RoboDK station: PICK1.rdk

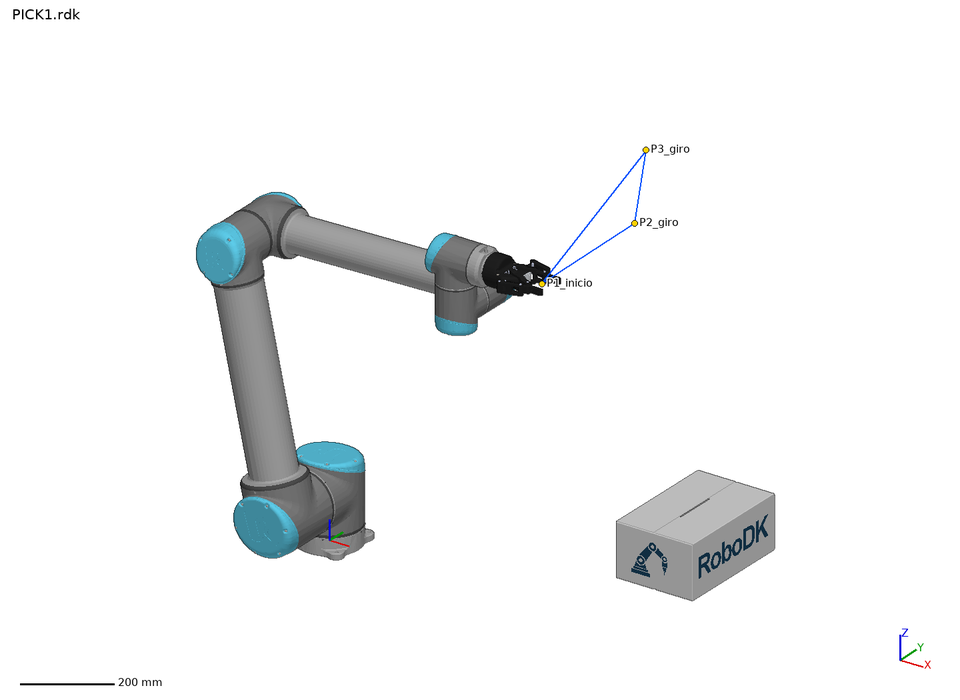
[picture v0: the station drawn from its stored meshes, robots at their saved joint values, targets as dots, program paths as lines]
Station Nueva Estación (1) (saved by RoboDK 6.1.1). Poses are relative to the parent item; angles as X-Y-Z fixed-axis rotations.
  - frame UR10 Base at (0, 0, 0) mm
    - robot UR10: 6 axes, payload 10 kg, reach 1300 mm, repeatability 0.1 mm, weight 28.9 kg
        modified DH rows (alpha deg, a mm, theta deg, d mm): 0, 0, 0, 128; 90, 0, 180, 0; 0, 612.7, 0, 0; 0, 571.6, 0, 163.9; -90, 0, 0, 115.7; 90, 0, 180, 92.2
        joint limits [-360, -360, -360, -360, -360, -360] to [360, 360, 360, 360, 360, 360]; home [0, -90, -90, 0, 90, 0]; saved at [0, -77.766, -100.839, -1.395, 90, 0]
      - tool RobotiQ 2F-85 Gripper (Closed), TCP at (0, 0, 130) mm, size 134.4 x 75 x 157.6 mm
    - target P1_inicio (Cartesian target) at (663.8, -163.9, 856.4) mm, rotated rx -90 ry 0 rz -90 deg; joints [0, -90, -90, 0, 90, 0] of UR10
    - target P2_giro (Cartesian target) at (656.82, 189.96, 856.4) mm, rotated rx -90 ry 0 rz -60 deg; joints [30, -90, -90, 0, 90, 0] of UR10
    - target P3_giro (Cartesian target) at (473.84, 492.92, 856.4) mm, rotated rx -90 ry 0 rz -30 deg; joints [60, -90, -90, 0, 90, 0] of UR10
    - object Caja at (600, 200, 0) mm, size 199 x 305.1 x 133.7 mm, geometry from Box-12x7in-Closed.sld
  - program Secuencia_UR10 (6 instructions, listed below)
  - Python program Prog2 (listed below)
  - Python program Prog3 (listed below)
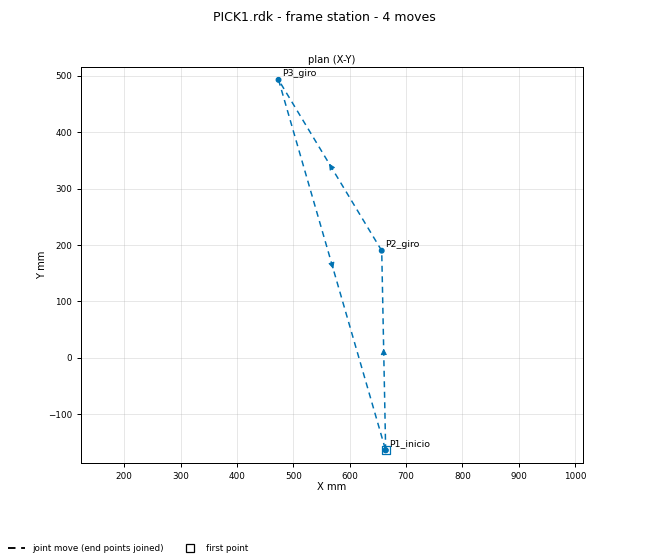
[picture p0: tool path of PICK1.rdk in frame station, 4 of 4 moves have a stored position in this frame; points joined in program order, loops and branches not executed]

--- program Secuencia_UR10 (robot UR10) ---
  Est. Ref.: UR10 Base
  MoveJ (P1_inicio)
  MoveJ (P2_giro)
  MoveJ (P3_giro)
  MoveJ (P1_inicio)
  Establecer velocidad (500.0 mm/s)

--- Python program Prog2 ---
from robodk.robolink import *

RDK = Robolink()

robot = RDK.Item('UR10', ITEM_TYPE_ROBOT)

p1 = RDK.Item('P1_inicio', ITEM_TYPE_TARGET)
p2 = RDK.Item('P2_giro', ITEM_TYPE_TARGET)
p3 = RDK.Item('P3_giro', ITEM_TYPE_TARGET)

# Verificar que existan los elementos
if not all(item.Valid() for item in [robot, p1, p2, p3]):
    raise Exception("No se encontro el robot o algun punto")

# Velocidad articular
robot.setSpeedJoints(20)

# Secuencia del brazo robotico
robot.MoveJ(p1)
robot.MoveJ(p2)
robot.MoveJ(p3)
robot.MoveJ(p1)

print("Secuencia completada")

--- Python program Prog3 ---
# -*- coding: utf-8 -*-
# Pick & Place UR10 + Robotiq 2F-85 en RoboDK (v2)
# La caja vuelve SIEMPRE a su origen al iniciar, asi se puede ejecutar muchas veces.

from robodk.robolink import *
from robodk.robomath import *

# ============ PARAMETROS (ajusta estos valores) ============
NOMBRE_ROBOT = 'UR10'
NOMBRE_CAJA = 'Caja'

# Posicion ORIGEN de la caja (respecto a la base del robot, mm)
ORIGEN_X, ORIGEN_Y, ORIGEN_Z = 600, -300, 0

# Desplazamiento del destino respecto al origen (mm, sistema de la base)
DESTINO_DX = 0
DESTINO_DY = 500
DESTINO_DZ = 0

ALTURA_SEGURA = 250     # mm sobre el punto de agarre (altura de viaje)
OFFSET_AGARRE_Z = 0     # mm: ajusta si la pinza queda muy alta/baja (+ sube, - baja)
ALTURA_CAJA = 0         # mm: sumar si el origen de la caja esta en su base

VEL_LINEAL = 150        # mm/s (bajada y subida lentas)
VEL_ARTICULAR = 60      # deg/s
# ===========================================================

RDK = Robolink()
robot = RDK.Item(NOMBRE_ROBOT, ITEM_TYPE_ROBOT)
caja = RDK.Item(NOMBRE_CAJA, ITEM_TYPE_OBJECT)

if not robot.Valid():
    raise Exception('No se encontro el robot "%s"' % NOMBRE_ROBOT)
if not caja.Valid():
    raise Exception('No se encontro el objeto "%s"' % NOMBRE_CAJA)

# Herramienta (la pinza Robotiq que cuelga del robot)
herramienta = RDK.Item('', ITEM_TYPE_TOOL)
for hijo in robot.Childs():
    if hijo.Type() == ITEM_TYPE_TOOL:
        herramienta = hijo
        break
if not herramienta.Valid():
    raise Exception('No se encontro la pinza (herramienta) en el robot')

base = robot.Parent()  # "UR10 Base"
robot.setPoseFrame(base)
robot.setPoseTool(herramienta)
robot.setSpeed(VEL_LINEAL, VEL_ARTICULAR)
robot.setRounding(5)

# --- Reiniciar la caja: soltarla de la pinza y devolverla al origen ---
herramienta.DetachAll(base)
caja.setParent(base)
caja.setPoseAbs(base.PoseAbs() * transl(ORIGEN_X, ORIGEN_Y, ORIGEN_Z))

# Posicion de la caja respecto a la base del robot
pose_caja = invH(base.PoseAbs()) * caja.PoseAbs()
x, y, z = pose_caja.Pos()

# Orientacion de la pinza: Z de la herramienta apuntando hacia abajo
ORIENTACION = rotx(pi)

z_agarre = z + ALTURA_CAJA + OFFSET_AGARRE_Z
pose_agarre = transl(x, y, z_agarre) * ORIENTACION
pose_sobre_caja = transl(x, y, z_agarre + ALTURA_SEGURA) * ORIENTACION

xd, yd, zd = x + DESTINO_DX, y + DESTINO_DY, z_agarre + DESTINO_DZ
pose_destino = transl(xd, yd, zd) * ORIENTACION
pose_sobre_destino = transl(xd, yd, zd + ALTURA_SEGURA) * ORIENTACION


def abrir_pinza():
    try:
        prog = RDK.Item('Gripper Open', ITEM_TYPE_PROGRAM)
        if prog.Valid():
            prog.RunProgram()
    except Exception:
        pass
    robot.RunInstruction('Abrir pinza', INSTRUCTION_COMMENT)
    pause(0.5)


def cerrar_pinza():
    try:
        prog = RDK.Item('Gripper Close', ITEM_TYPE_PROGRAM)
        if prog.Valid():
            prog.RunProgram()
    except Exception:
        pass
    robot.RunInstruction('Cerrar pinza', INSTRUCTION_COMMENT)
    pause(0.5)


# Comprobacion de alcance antes de moverse
for nombre, p in [('sobre caja', pose_sobre_caja), ('agarre', pose_agarre),
                  ('sobre destino', pose_sobre_destino), ('destino', pose_destino)]:
    joints = robot.SolveIK(p)
    if len(joints.list()) < 6:
        raise Exception('Posicion "%s" fuera de alcance. Cambia ORIGEN/DESTINO o la altura.' % nombre)

# ===================== SECUENCIA =====================
robot.RunInstruction('Inicio pick and place', INSTRUCTION_COMMENT)

# 1) Ir a la posicion de inicio (si existe el target P1_inicio)
inicio = RDK.Item('P1_inicio', ITEM_TYPE_TARGET)
if inicio.Valid():
    robot.MoveJ(inicio)

# 2) Abrir pinza y colocarse sobre la caja
abrir_pinza()
robot.MoveJ(pose_sobre_caja)

# 3) Agacharse hasta la caja (movimiento lineal, lento)
robot.MoveL(pose_agarre)

# 4) Cerrar pinza y agarrar la caja
cerrar_pinza()
herramienta.AttachClosest()

# 5) Levantar la caja
robot.MoveL(pose_sobre_caja)

# 6) Transportar hasta sobre el destino
robot.MoveJ(pose_sobre_destino)

# 7) Agacharse para dejar la caja
robot.MoveL(pose_destino)

# 8) Soltar la caja y abrir pinza
herramienta.DetachAll(base)
abrir_pinza()

# 9) Subir y volver a inicio
robot.MoveL(pose_sobre_destino)
if inicio.Valid():
    robot.MoveJ(inicio)

robot.RunInstruction('Fin pick and place', INSTRUCTION_COMMENT)
print('Listo: la caja fue movida.')
